(* IEC 61131-3 sources: machine-design-framework/examples/pick-glue-place/plc/targets/sim, 2 files *)

(* ---- GVL_Sim.st ---- *)
(* SIL-only globals written by the plant model. Not part of any real target. *)
VAR_GLOBAL
    xSimDriveFaultX : BOOL;
    xSimDriveFaultZ : BOOL;
END_VAR

(* ---- FB_Axis.st ---- *)
(* SIL implementation of FB_Axis: the plant model stands in for drive and motion. *)
FUNCTION_BLOCK FB_Axis
VAR_INPUT
    xEnable  : BOOL;
    xSimFault: BOOL;     (* set by the SIL plant to inject a drive fault *)
END_VAR
VAR_OUTPUT
    xReady   : BOOL;
    xError   : BOOL;
    iErrorId : INT;
END_VAR
xError := xSimFault;
IF xError THEN
    iErrorId := 9001;
ELSE
    iErrorId := 0;
END_IF;
xReady := xEnable AND NOT xError;
END_FUNCTION_BLOCK
